(* IEC 61131-3 sources: rusty/compiler/plc_cfc/fixtures/blocks/valid/action_program, 1 file *)

(* ---- P.st ---- *)
PROGRAM P
VAR_INPUT
    step : DINT;
END_VAR
VAR_OUTPUT
    out : DINT;
END_VAR
END_PROGRAM

ACTIONS
    ACTION bump
        out := out + step;
    END_ACTION
END_ACTIONS
